Fanuc KAREL source: KT00275.KL

PROGRAM KT00275
%NOLOCKGROUP
VAR
  P1: POSITION
  P2: POSITION
  OUT: BOOLEAN
BEGIN
  OUT = P1 = P2
END KT00275
